Staubli VAL3: refreshData.pgx

program refreshData(num x_nIndex)
  local tool l_tTool
begin
  nFrame[0]=safeTemp:zZoneItem[x_nIndex].fBase.trsf.x
  nFrame[1]=safeTemp:zZoneItem[x_nIndex].fBase.trsf.y
  nFrame[2]=safeTemp:zZoneItem[x_nIndex].fBase.trsf.z
  nFrame[3]=safeTemp:zZoneItem[x_nIndex].fBase.trsf.rx
  nFrame[4]=safeTemp:zZoneItem[x_nIndex].fBase.trsf.ry
  nFrame[5]=safeTemp:zZoneItem[x_nIndex].fBase.trsf.rz
  fFrame.trsf=safeTemp:zZoneItem[x_nIndex].fBase.trsf
  call saveData:getTool(saveData:nJogTool,tTool)
  $jogContext(tTool,fFrame,0)

  nTRSF1[0]=safeTemp:zZoneItem[x_nIndex].pFirst.trsf.x
  nTRSF1[1]=safeTemp:zZoneItem[x_nIndex].pFirst.trsf.y
  nTRSF1[2]=safeTemp:zZoneItem[x_nIndex].pFirst.trsf.z
  nTRSF1[3]=safeTemp:zZoneItem[x_nIndex].pFirst.trsf.rx
  nTRSF1[4]=safeTemp:zZoneItem[x_nIndex].pFirst.trsf.ry
  nTRSF1[5]=safeTemp:zZoneItem[x_nIndex].pFirst.trsf.rz

  nTRSF2[0]=safeTemp:zZoneItem[x_nIndex].pSecond.trsf.x
  nTRSF2[1]=safeTemp:zZoneItem[x_nIndex].pSecond.trsf.y
  nTRSF2[2]=safeTemp:zZoneItem[x_nIndex].pSecond.trsf.z
  nTRSF2[3]=safeTemp:zZoneItem[x_nIndex].pSecond.trsf.rx
  nTRSF2[4]=safeTemp:zZoneItem[x_nIndex].pSecond.trsf.ry
  nTRSF2[5]=safeTemp:zZoneItem[x_nIndex].pSecond.trsf.rz

  sComment=safeTemp:zZoneItem[x_nIndex].sID

end
